Fanuc KAREL source: KT00129.KL

PROGRAM KT00129
%NOLOCKGROUP
VAR
  I1: INTEGER
  I2: INTEGER
  OUT: INTEGER
BEGIN
  I1 = 2
  I2 = 3
  I1 = 2
  I2 = 3
  OUT = I1 DIV I2
END KT00129
